Staubli VAL3: Motion.dtx

public mdesc mNomSpeed = {accel=25, vel=20, decel=25, blend=off, leave=0, reach=0}
public mdesc mFine = {accel=10, vel=10, decel=10, blend=off, leave=0, reach=0}
public joint jHome
public tool tTool = {fatherId=flange[0]}
